// Mitsubishi GX Works2 project: 1127シーケンサ特殊命令など使用して改良   PLC: FX3G

PROGRAM MAIN
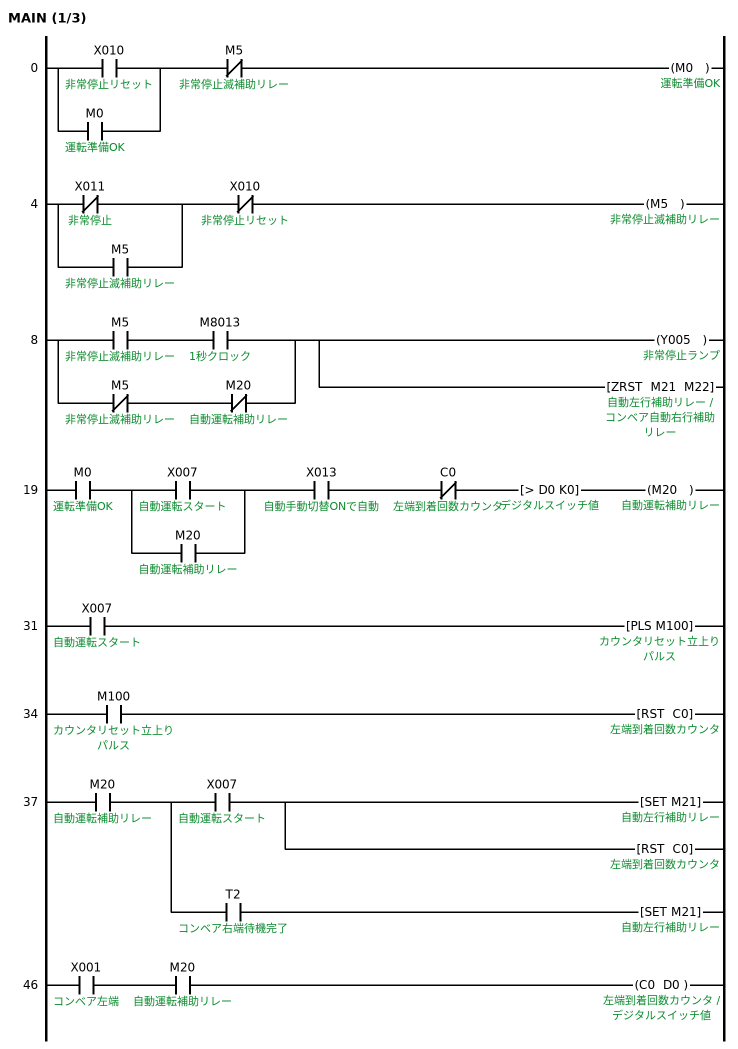
0     LD      X010  ; 非常停止リセット
      OR      M0  ; 運転準備OK
      ANI     M5  ; 非常停止滅補助リレー
      OUT     M0  ; 運転準備OK
4     LDI     X011  ; 非常停止
      OR      M5  ; 非常停止滅補助リレー
      ANI     X010  ; 非常停止リセット
      OUT     M5  ; 非常停止滅補助リレー
8     LD      M5  ; 非常停止滅補助リレー
      AND     M8013  ; 1秒クロック
      LDI     M5  ; 非常停止滅補助リレー
      ANI     M20  ; 自動運転補助リレー
      ORB
      OUT     Y005  ; 非常停止ランプ
      ZRST    M21 M22  ; 自動左行補助リレー / コンベア自動右行補助リレー
19    LD      M0  ; 運転準備OK
      LD      X007  ; 自動運転スタート
      OR      M20  ; 自動運転補助リレー
      ANB
      AND     X013  ; 自動手動切替ONで自動
      ANI     C0  ; 左端到着回数カウンタ
      AND>    D0 K0  ; デジタルスイッチ値
      OUT     M20  ; 自動運転補助リレー
31    LD      X007  ; 自動運転スタート
      PLS     M100  ; カウンタリセット立上りパルス
34    LD      M100  ; カウンタリセット立上りパルス
      RST     C0  ; 左端到着回数カウンタ
37    LD      M20  ; 自動運転補助リレー
      MPS
      AND     X007  ; 自動運転スタート
      SET     M21  ; 自動左行補助リレー
      RST     C0  ; 左端到着回数カウンタ
      MPP
      AND     T2  ; コンベア右端待機完了
      SET     M21  ; 自動左行補助リレー
46    LD      X001  ; コンベア左端
      AND     M20  ; 自動運転補助リレー
      OUT     C0 D0  ; 左端到着回数カウンタ / デジタルスイッチ値
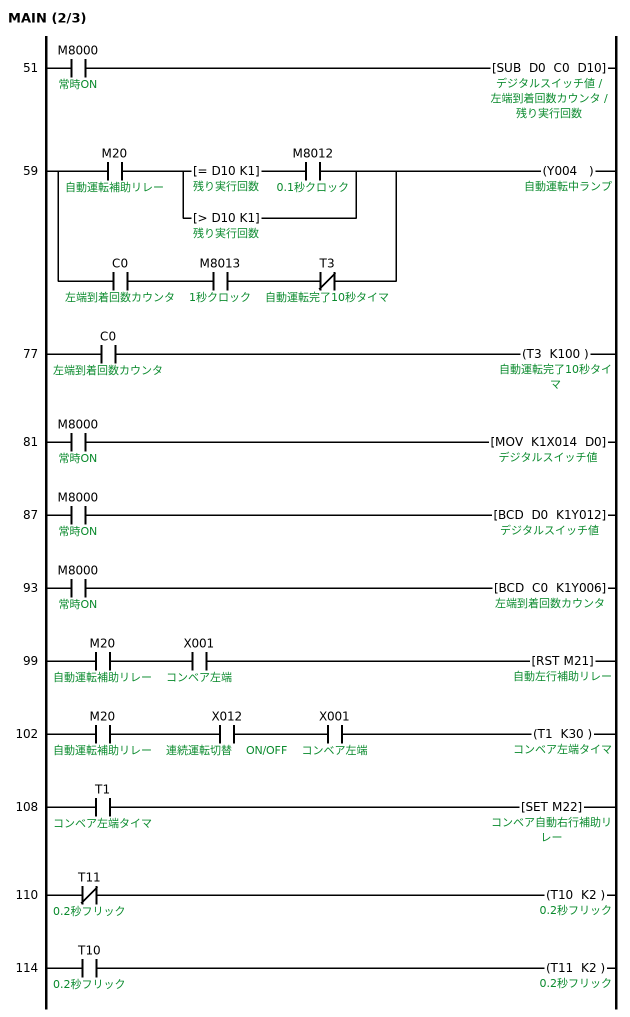
51    LD      M8000  ; 常時ON
      SUB     D0 C0 D10  ; 残り実行回数
59    LD      M20  ; 自動運転補助リレー
      LD=     D10 K1  ; 残り実行回数
      AND     M8012  ; 0.1秒クロック
      OR>     D10 K1  ; 残り実行回数
      ANB
      LD      C0  ; 左端到着回数カウンタ
      AND     M8013  ; 1秒クロック
      ANI     T3  ; 自動運転完了10秒タイマ
      ORB
      OUT     Y004  ; 自動運転中ランプ
77    LD      C0  ; 左端到着回数カウンタ
      OUT     T3 K100  ; 自動運転完了10秒タイマ
81    LD      M8000  ; 常時ON
      MOV     K1X014 D0  ; デジタルスイッチ入力値転送
87    LD      M8000  ; 常時ON
      BCD     D0 K1Y012
93    LD      M8000  ; 常時ON
      BCD     C0 K1Y006
99    LD      M20  ; 自動運転補助リレー
      AND     X001  ; コンベア左端
      RST     M21  ; 自動左行補助リレー
102   LD      M20  ; 自動運転補助リレー
      AND     X012  ; 連続運転切替    ON/OFF
      AND     X001  ; コンベア左端
      OUT     T1 K30  ; コンベア左端タイマ
108   LD      T1  ; コンベア左端タイマ
      SET     M22  ; コンベア自動右行補助リレー
110   LDI     T11  ; 0.2秒フリック
      OUT     T10 K2  ; 0.2秒フリック
114   LD      T10  ; 0.2秒フリック
      OUT     T11 K2  ; 0.2秒フリック
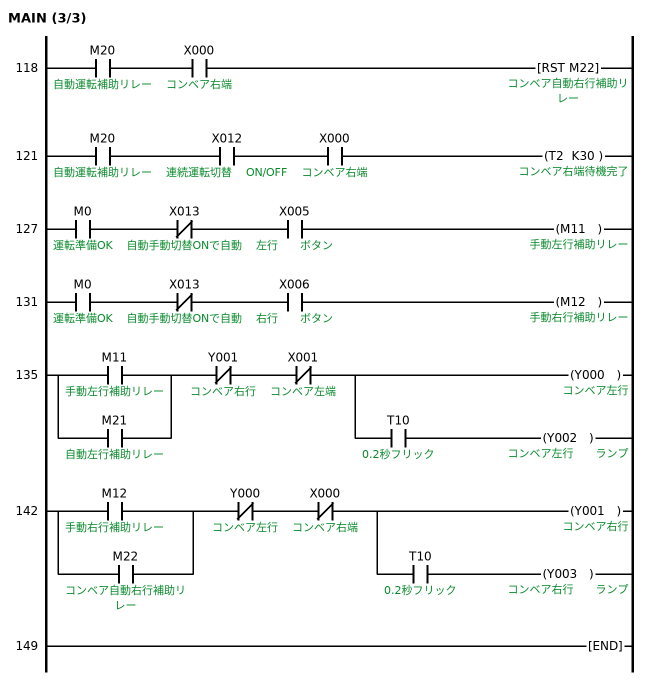
118   LD      M20  ; 自動運転補助リレー
      AND     X000  ; コンベア右端
      RST     M22  ; コンベア自動右行補助リレー
121   LD      M20  ; 自動運転補助リレー
      AND     X012  ; 連続運転切替    ON/OFF
      AND     X000  ; コンベア右端
      OUT     T2 K30  ; コンベア右端待機完了
127   LD      M0  ; 運転準備OK
      ANI     X013  ; 自動手動切替ONで自動
      AND     X005  ; 左行　　ボタン
      OUT     M11  ; 手動左行補助リレー
131   LD      M0  ; 運転準備OK
      ANI     X013  ; 自動手動切替ONで自動
      AND     X006  ; 右行　　ボタン
      OUT     M12  ; 手動右行補助リレー
135   LD      M11  ; 手動左行補助リレー
      OR      M21  ; 自動左行補助リレー
      ANI     Y001  ; コンベア右行
      ANI     X001  ; コンベア左端
      OUT     Y000  ; コンベア左行
      AND     T10  ; 0.2秒フリック
      OUT     Y002  ; コンベア左行　　ランプ
142   LD      M12  ; 手動右行補助リレー
      OR      M22  ; コンベア自動右行補助リレー
      ANI     Y000  ; コンベア左行
      ANI     X000  ; コンベア右端
      OUT     Y001  ; コンベア右行
      AND     T10  ; 0.2秒フリック
      OUT     Y003  ; コンベア右行　　ランプ
149   END
END_PROGRAM

// device comments not shown above
Y030  ; 7セグ表示
M55  ; 非常停止ランプ　補助リレー
T44  ; 非常停止ランプ点滅タイマOFF
T55  ; 非常停止ランプ点滅タイマON
